TYPE ST_CIP_Request :
STRUCT
	eType	: E_CIP_Type;
	eClient	: E_CIP_Usage;
	nClientId	: INT;					//1..30, 0 for eLocal
	eClientType	: E_Anybus_ClientType;	//eExternal only
	eStartState	: E_Element_State_Long;	//eExternal only: first stage, by the GAD wash type

END_STRUCT
END_TYPE

(* stored: Version 1.1.0.1, ProductVersion 3.1.4024.12
   DUT ST_CIP_Request: Id {9bd869e0-a3c9-4647-8549-556577cea663} *)
